(* IEC 61131-3 sources: plcassist-cli/packages/volt-lsp-iec/test-corpus/bakon-nano/Device/Plc Logic/Application/Library Manager/L_SMHP_ModuleHandler, 20 files *)

(* ---- CONDITIONALSHOW_WHITELIST_LOG.gvl ---- *)
VAR_GLOBAL
END_VAR

(* ---- GETBOOLEANPROPERTY.fun ---- *)
FUNCTION GETBOOLEANPROPERTY : BOOL
VAR_INPUT
	STKEY : WSTRING;
END_VAR
END_FUNCTION

(* ---- GETCOMPANY.fun ---- *)
FUNCTION GETCOMPANY : WSTRING
END_FUNCTION

(* ---- GETNUMBERPROPERTY.fun ---- *)
FUNCTION GETNUMBERPROPERTY : DINT
VAR_INPUT
	STKEY : WSTRING;
END_VAR
END_FUNCTION

(* ---- GETTEXTPROPERTY.fun ---- *)
FUNCTION GETTEXTPROPERTY : WSTRING
VAR_INPUT
	STKEY : WSTRING;
END_VAR
END_FUNCTION

(* ---- GETTEXTPROPERTY2.fun ---- *)
FUNCTION GETTEXTPROPERTY2 : POINTER TO WSTRING
VAR_INPUT
	STKEY : WSTRING;
END_VAR
END_FUNCTION

(* ---- GETTITLE.fun ---- *)
FUNCTION GETTITLE : WSTRING
END_FUNCTION

(* ---- GETVERSION.fun ---- *)
FUNCTION GETVERSION : VERSION
END_FUNCTION

(* ---- GETVERSIONPROPERTY.fun ---- *)
FUNCTION GETVERSIONPROPERTY : VERSION
VAR_INPUT
	STKEY : WSTRING;
END_VAR
END_FUNCTION

(* ---- L_SMHP_CALLSERVICEFUNCTION.fun ---- *)
FUNCTION L_SMHP_CALLSERVICEFUNCTION : UDINT
VAR_INPUT
	MODULEHANDLE : RTS_IEC_HANDLE;
	SERVICEID : DWORD;
	COMMANDID : DWORD;
	SZDATA : UDINT;
	PDATA : POINTER TO BYTE;
END_VAR
END_FUNCTION

(* ---- L_SMHP_CONFIGURESERVICE.fun ---- *)
FUNCTION L_SMHP_CONFIGURESERVICE : UDINT
VAR_INPUT
	SERVICEID : DWORD;
	COMMANDID : DWORD;
	SZDATA : UDINT;
	PDATA : POINTER TO BYTE;
END_VAR
END_FUNCTION

(* ---- L_SMHP_CONFIGURESERVICEAVAILABLE.fun ---- *)
FUNCTION L_SMHP_CONFIGURESERVICEAVAILABLE : BOOL
VAR_INPUT
	SERVICEID : DWORD;
	COMMANDID : DWORD;
END_VAR
END_FUNCTION

(* ---- L_SMHP_GETAVAILABLESERVICES.fun ---- *)
FUNCTION L_SMHP_GETAVAILABLESERVICES : UDINT
VAR_INPUT
	SZREQUESTEDSERVICES : UDINT;
	PREQUESTEDSERVICE : POINTER TO BYTE;
END_VAR
END_FUNCTION

(* ---- L_SMHP_REGISTERCOMPONENT.fun ---- *)
FUNCTION L_SMHP_REGISTERCOMPONENT : RTS_IEC_HANDLE
VAR_INPUT
	COMPTYPE : DWORD;
	LAYER : BYTE;
	XACTIVE : BOOL;
	SCOMPONENTNAME : POINTER TO STRING;
	SINSTANCEPATH : POINTER TO STRING;
	SZREQUESTEDSERVICE : UDINT;
	PREQUESTEDSERVICE : POINTER TO BYTE;
END_VAR
END_FUNCTION

(* ---- L_SMHP_REGISTERCOMPONENT_V2.fun ---- *)
FUNCTION L_SMHP_REGISTERCOMPONENT_V2 : RTS_IEC_HANDLE
VAR_INPUT
	COMPTYPE : DWORD;
	COMPSUBTYPE : DWORD;
	LAYER : BYTE;
	XACTIVE : BOOL;
	SCOMPONENTNAME : POINTER TO STRING;
	SINSTANCEPATH : POINTER TO STRING;
	SZREQUESTEDSERVICE : UDINT;
	PREQUESTEDSERVICE : POINTER TO BYTE;
END_VAR
END_FUNCTION

(* ---- L_SMHP_SERVICEFUNCTIONAVAILABLE.fun ---- *)
FUNCTION L_SMHP_SERVICEFUNCTIONAVAILABLE : BOOL
VAR_INPUT
	SERVICEID : DWORD;
	COMMANDID : DWORD;
END_VAR
END_FUNCTION

(* ---- L_SMHP_UNREGISTERCOMPONENT.fun ---- *)
FUNCTION L_SMHP_UNREGISTERCOMPONENT : UDINT
VAR_INPUT
	MODULEHANDLE : RTS_IEC_HANDLE;
END_VAR
END_FUNCTION

(* ---- L_SMHP_UPDATECOMPONENTINFO.fun ---- *)
FUNCTION L_SMHP_UPDATECOMPONENTINFO : UDINT
VAR_INPUT
	MODULEHANDLE : RTS_IEC_HANDLE;
	COMMANDID : DWORD;
	SZDATA : UDINT;
	PDATA : POINTER TO BYTE;
END_VAR
END_FUNCTION

(* ---- L_SMHP_UPDATESERVICEINFO.fun ---- *)
FUNCTION L_SMHP_UPDATESERVICEINFO : UDINT
VAR_INPUT
	MODULEHANDLE : RTS_IEC_HANDLE;
	SZREQUESTEDSERVICE : UDINT;
	PREQUESTEDSERVICE : POINTER TO BYTE;
END_VAR
END_FUNCTION

(* ---- L_SMHP_WRITECOMPONENTLIST.fun ---- *)
FUNCTION L_SMHP_WRITECOMPONENTLIST : UDINT
VAR_INPUT
	PFILENAME : POINTER TO STRING;
END_VAR
END_FUNCTION
